DATA_BLOCK "EC_Positioning_DB"
{ S7_Optimized_Access := 'FALSE' }
VERSION : 0.1
NON_RETAIN
"EC_Positioning"
BEGIN
END_DATA_BLOCK

